(* IEC 61131-3 sources: plc-iiot-stack/src/POUs/Iiot/F_IiotAlarmReasonText, 2 files *)

(* ---- F_IiotAlarmReasonText.decl.st ---- *)
// Назначение: имя причины события тревоги для поля reason.
// Автор:      kr0nsch
// Версия:     0.1.0
// Документ:   docs/plc_mqtt.md, раздел «Тревоги»
FUNCTION F_IiotAlarmReasonText : STRING(GVL_Const.IIOT_TEXT_LEN)
VAR_INPUT
    eReason : E_IiotAlarmReason;
END_VAR

(* ---- F_IiotAlarmReasonText.impl.st ---- *)
CASE eReason OF
    E_IiotAlarmReason.Activated:
        F_IiotAlarmReasonText := 'Activated';
    E_IiotAlarmReason.Cleared:
        F_IiotAlarmReasonText := 'Cleared';
    E_IiotAlarmReason.Acked:
        F_IiotAlarmReasonText := 'Acked';
    E_IiotAlarmReason.Shelved:
        F_IiotAlarmReasonText := 'Shelved';
    E_IiotAlarmReason.Unshelved:
        F_IiotAlarmReasonText := 'Unshelved';
    E_IiotAlarmReason.ShelveExpired:
        F_IiotAlarmReasonText := 'ShelveExpired';
    E_IiotAlarmReason.Suppressed:
        F_IiotAlarmReasonText := 'Suppressed';
    E_IiotAlarmReason.Unsuppressed:
        F_IiotAlarmReasonText := 'Unsuppressed';
    E_IiotAlarmReason.OosOn:
        F_IiotAlarmReasonText := 'OosOn';
ELSE
    F_IiotAlarmReasonText := 'OosOff';
END_CASE
